Fanuc KAREL source: kd00051.KL

-- PROVISIONAL review KL for V1013-1; original PC SHA256 6ffc7c6f7322692f010cd36729554ed56665b5a549f5756baba35c0fe20ec65e
-- Incomplete behavior may be omitted. Consult companion uncertainty JSON. Do not deploy.
PROGRAM KD00051
%NOLOCKGROUP
VAR
  I : INTEGER
  J : INTEGER
  B : BOOLEAN
  R : REAL
  S : STRING[80]
-- UNRESOLVED_DECL P type=000101
BEGIN
  -- UNRESOLVED_PC offsets 5-30; opcodes 01,22,1C,2E,0A,82,0B
  -- UNRESOLVED_PC offsets 35-39; opcodes 7F
END KD00051
